// SIMATIC S7-200 project (STEP 7-Micro/WIN), CPU 224 CN REL 02.01

SYMBOL_TABLE 用户定义1
允许加工             V1000.6
停止               M0.1
准备就绪             M0.0
全线模式             V1010.1
网络正常             V1010.0
加工完成             V1010.2
物料台物料检测          I0.0
料台夹紧检测           I0.1
料台伸出到位检测         I0.2
料台缩回到位检测         I0.3
加工压头上限检测         I0.4
加工压头下限检测         I0.5
停止按钮             I1.2
启动按钮             I1.3
急停按钮             I1.4
单机全线             I1.5
夹紧电磁阀            Q0.0
料台伸缩电磁阀          Q0.2
加工压头电磁阀          Q0.3
正常工作指示           Q0.7
设备运行指示           Q1.0
红色指示灯            Q1.1
END_SYMBOL_TABLE

ORGANIZATION_BLOCK 主程序:OB1
TITLE=程序注释
BEGIN
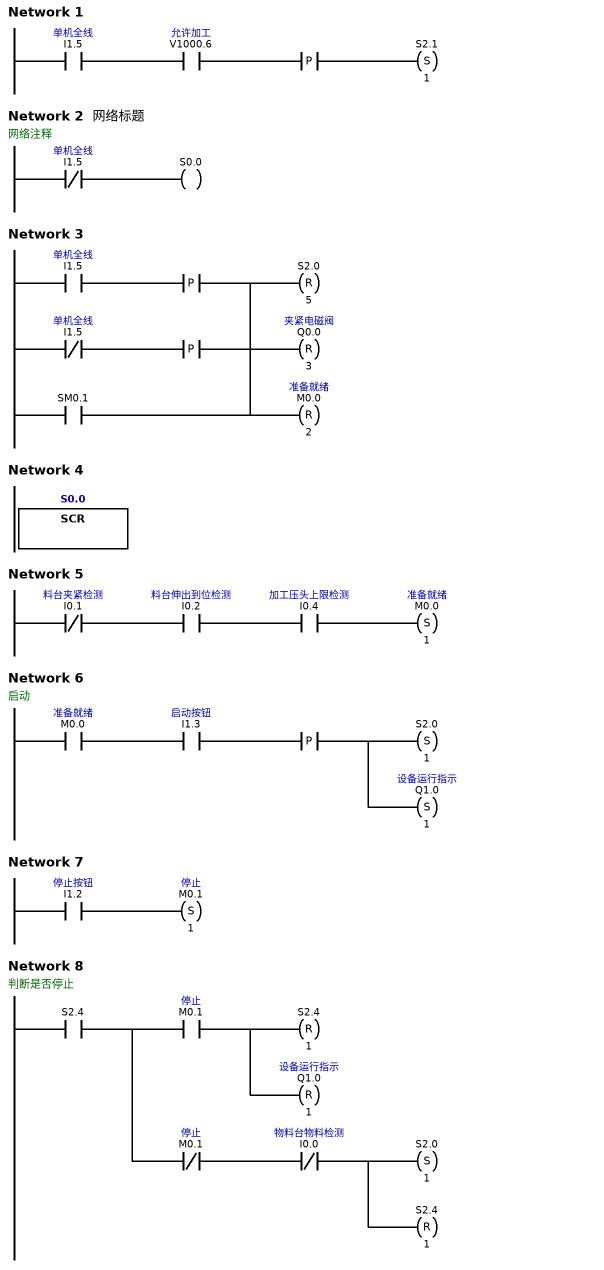
Network 1
LD     单机全线:I1.5
A      允许加工:V1000.6
EU
S      S2.1, 1
Network 2 // 网络标题
// 网络注释
LDN    单机全线:I1.5
=      S0.0
Network 3
LD     单机全线:I1.5
EU
LDN    单机全线:I1.5
EU
OLD
O      SM0.1
R      S2.0, 5
R      夹紧电磁阀:Q0.0, 3
R      准备就绪:M0.0, 2
Network 4
LSCR   S0.0
Network 5
LDN    料台夹紧检测:I0.1
A      料台伸出到位检测:I0.2
A      加工压头上限检测:I0.4
S      准备就绪:M0.0, 1
Network 6
// 启动
LD     准备就绪:M0.0
A      启动按钮:I1.3
EU
S      S2.0, 1
S      设备运行指示:Q1.0, 1
Network 7
LD     停止按钮:I1.2
S      停止:M0.1, 1
Network 8
// 判断是否停止
LD     S2.4
LPS
A      停止:M0.1
R      S2.4, 1
R      设备运行指示:Q1.0, 1
LPP
AN     停止:M0.1
AN     物料台物料检测:I0.0
S      S2.0, 1
R      S2.4, 1
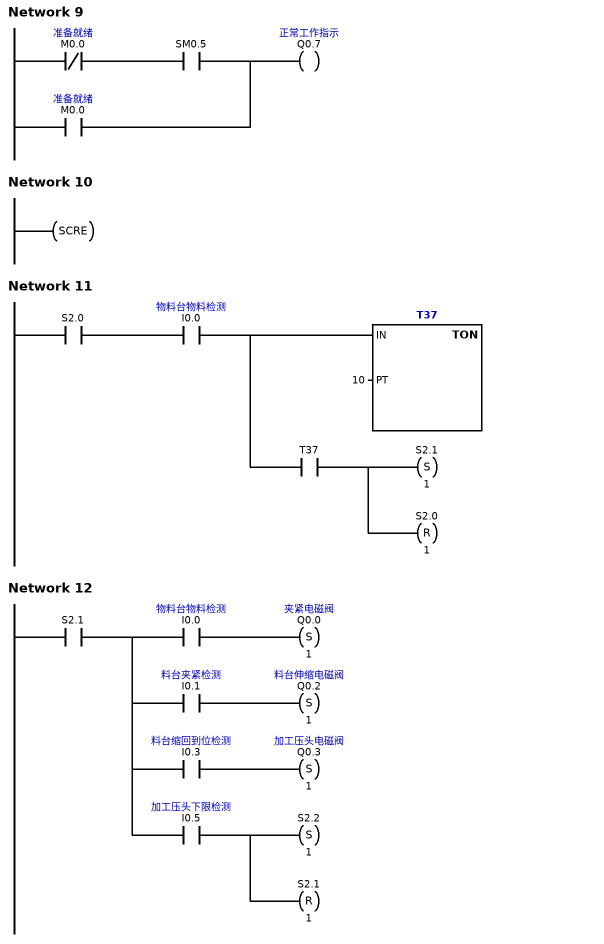
Network 9
LDN    准备就绪:M0.0
A      SM0.5
O      准备就绪:M0.0
=      正常工作指示:Q0.7
Network 10
SCRE
Network 11
LD     S2.0
A      物料台物料检测:I0.0
TON    T37, 10
A      T37
S      S2.1, 1
R      S2.0, 1
Network 12
LD     S2.1
LPS
A      物料台物料检测:I0.0
S      夹紧电磁阀:Q0.0, 1
LRD
A      料台夹紧检测:I0.1
S      料台伸缩电磁阀:Q0.2, 1
LRD
A      料台缩回到位检测:I0.3
S      加工压头电磁阀:Q0.3, 1
LPP
A      加工压头下限检测:I0.5
S      S2.2, 1
R      S2.1, 1
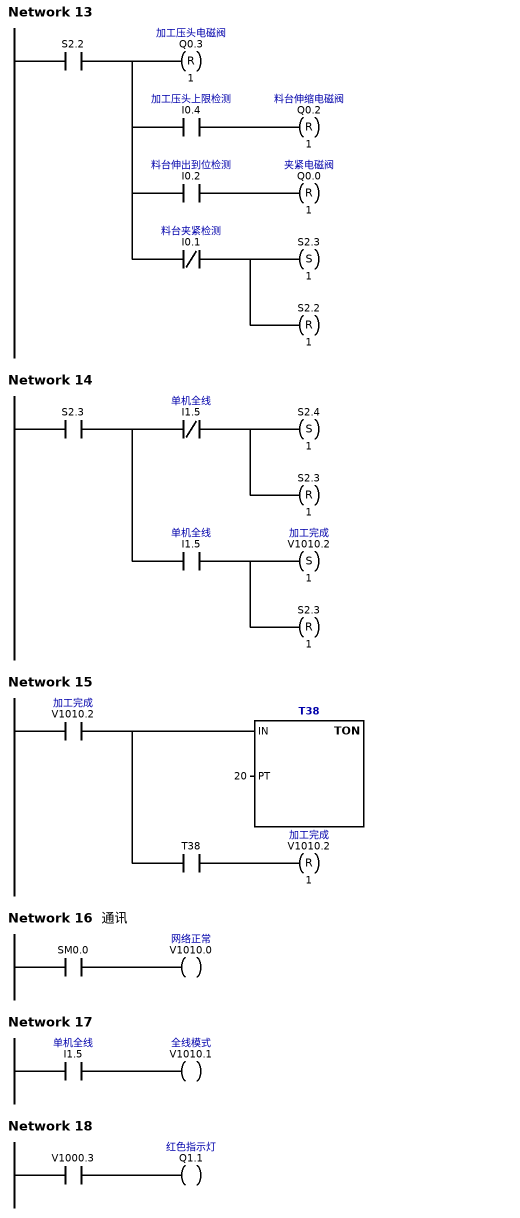
Network 13
LD     S2.2
LPS
R      加工压头电磁阀:Q0.3, 1
A      加工压头上限检测:I0.4
R      料台伸缩电磁阀:Q0.2, 1
LRD
A      料台伸出到位检测:I0.2
R      夹紧电磁阀:Q0.0, 1
LPP
AN     料台夹紧检测:I0.1
S      S2.3, 1
R      S2.2, 1
Network 14
LD     S2.3
LPS
AN     单机全线:I1.5
S      S2.4, 1
R      S2.3, 1
LPP
A      单机全线:I1.5
S      加工完成:V1010.2, 1
R      S2.3, 1
Network 15
LD     加工完成:V1010.2
TON    T38, 20
A      T38
R      加工完成:V1010.2, 1
Network 16 // 通讯
LD     SM0.0
=      网络正常:V1010.0
Network 17
LD     单机全线:I1.5
=      全线模式:V1010.1
Network 18
LD     V1000.3
=      红色指示灯:Q1.1
END_ORGANIZATION_BLOCK
